// TIA Portal V19 export
DATA_BLOCK "Tacho2_EM04"   // DB5
VERSION : 1.0
// stored: InstanceOfName EM04_Insumos, InstanceOfType FB
"EM04_Insumos"
   // VAR_INPUT
   //    In : "EM04_Input";
   //    LevelPV : Real;
   // END_VAR
   // VAR_OUTPUT
   //    Out : "EM04_Output";
   //    CM_Vlv_Cristal_Out : Array[1..3] of Bool;
   //    TimeoutAlarm : Bool;
   //    SensorAlarm : Bool;
   //    CMAlarm : Bool;
   // END_VAR
   // VAR
   //    State : Int;
   //    ActiveAction : Int;
   //    ActiveValveIndex : Int;
   //    ElapsedPrev : Time;
   //    InjectionDone : Bool;
   //    AlarmLatched : Bool;
   //    FaultCode : Int;
   //    TimerInjection { S7_SetPoint := 'True'} : TON_TIME;
   //    TimerLevel { S7_SetPoint := 'True'} : TON_TIME;
   //    TimerTimeout { S7_SetPoint := 'True'} : TON_TIME;
   //    TrigStart { S7_SetPoint := 'True'} : R_TRIG;
   //    TrigStop { S7_SetPoint := 'True'} : R_TRIG;
   //    TrigHold { S7_SetPoint := 'True'} : R_TRIG;
   //    TrigAbort { S7_SetPoint := 'True'} : R_TRIG;
   //    TrigReset { S7_SetPoint := 'True'} : R_TRIG;
   //    CM_Vlv_Cristal { S7_SetPoint := 'True'} : Array[1..3] of "VlvL";
   // END_VAR
BEGIN
   In.TargetLevelSP := 50.0;
END_DATA_BLOCK
